Fanuc KAREL source: KT00978.KL

PROGRAM KT00978
%NOLOCKGROUP
VAR
  ENTRY: INTEGER
  PNAME: STRING[80]
  VNAME: STRING[80]
  STATUS: INTEGER
  VALUE: QUEUE_TYPE
BEGIN
  ENTRY = 0
  PNAME = ''
  VNAME = 'VALUE'
  SET_VAR(ENTRY, PNAME, VNAME, VALUE, STATUS)
END KT00978
